Fanuc KAREL source: ka00011.KL

-- PROVISIONAL review KL for V1013-1; original PC SHA256 7360e904d2c7ee1dd1bdd7d99eec25b3356701c621d0a9ac087e83b6fbc24066
-- Incomplete behavior may be omitted. Consult companion uncertainty JSON. Do not deploy.
PROGRAM KA00011
%NOLOCKGROUP
VAR
  SRC : INTEGER
-- UNRESOLVED_DECL DST type=002018
BEGIN
  -- UNRESOLVED_PC offsets 5-16; opcodes 2E,23
  -- UNRESOLVED_PC offsets 21-36; opcodes 21,22,9D,33,B2
  -- UNRESOLVED_PC offsets 41-45; opcodes 7F
END KA00011
